// TIA Portal V21 export
DATA_BLOCK "IDB_Mixed"   // DB23
// stored: InstanceOfName FB_Mixed, InstanceOfType FB
"FB_Mixed"
   // VAR_INPUT
   //    Start : Bool;
   //    RawValue : Int;
   // END_VAR
   // VAR_OUTPUT
   //    Running : Bool;
   //    Scaled : Real;
   //    AboveLimit : Bool;
   // END_VAR
   // VAR
   //    Factor : Real;
   //    Limit : Real;
   //    IsAbove : Bool;
   // END_VAR
BEGIN
END_DATA_BLOCK
